Fanuc KAREL source: kt00368.KL

-- PROVISIONAL review KL for V770-1; original PC SHA256 f05b54c1fad7ee41a159d6945e12ff9f3f7bcb8a83502d5e91fc5c98016d5678
-- Incomplete behavior may be omitted. Consult companion uncertainty JSON. Do not deploy.
PROGRAM KT00368
%NOLOCKGROUP
VAR
  I1 : INTEGER
  OUT : BOOLEAN
-- UNRESOLVED_DECL H2 type=002017
BEGIN
  -- UNRESOLVED_PC offsets 5-16; opcodes 2E,23
  -- UNRESOLVED_PC offsets 21-35; opcodes 2E,22,9D,33,B4
  -- UNRESOLVED_PC offsets 40-62; opcodes 21,22,9D,33,B3,5A,23
  -- UNRESOLVED_PC offsets 67-71; opcodes 7F
END KT00368
